{attribute 'qualified_only'}
{attribute 'strict'}
TYPE E_CmControlModuleCmd :
(
	NoCmd
);
END_TYPE

(* stored: Version 1.1.0.1, ProductVersion 3.1.4024.12
   DUT E_CmControlModuleCmd: Id {0fb8c39d-988c-4731-b3e3-d628f8bc00c4} *)
